FUNCTION_BLOCK FB_Light
VAR_INPUT
	bToggle : BOOL;
	bSetValid : BOOL;
	bTargetOn : BOOL;
END_VAR
VAR_OUTPUT
	bOn : BOOL;
END_VAR

IF bToggle THEN
	bOn := NOT bOn;
ELSIF bSetValid THEN
	bOn := bTargetOn;
END_IF

END_FUNCTION_BLOCK

(* stored: Version 1.1.0.1
   POU FB_Light: Id {40bd1988-e0d2-44ea-a579-af0915fd1114}, SpecialFunc None *)
